Fanuc KAREL source: kt00012.KL

-- PROVISIONAL review KL for V1013-1; original PC SHA256 02a34bf66193e1de4c26670054779a039fbb2b6cfb32eb01d97544c0d50c97d2
-- Incomplete behavior may be omitted. Consult companion uncertainty JSON. Do not deploy.
PROGRAM KT00012
%NOLOCKGROUP
VAR
  R1 : REAL
  R2 : REAL
  OUT : REAL
BEGIN
  -- UNRESOLVED_PC offsets 5-16; opcodes 2E,23
  -- UNRESOLVED_PC offsets 21-32; opcodes 2E,23
  -- UNRESOLVED_PC offsets 37-48; opcodes 2E,23
  -- UNRESOLVED_PC offsets 53-64; opcodes 2E,23
  -- UNRESOLVED_PC offsets 69-88; opcodes 21,21,69,23
  -- UNRESOLVED_PC offsets 93-97; opcodes 7F
END KT00012
